// TIA Portal project "FactoryIO_Template_S7-1200_V15_V16" (V16)
// Vorlageprojekt für das Buch mit Zielsystem S7-1200

(* hardware
DEVICE "S7-1200-Station_1"  S7-1200 Station
   slot 0: "Baugruppenträger_0"  Rack  V1.0
   slot 1: "PLC_1"  CPU 1212C AC/DC/Rly  6ES7 212-1BE40-0XB0  V4.4
DEVICE "HMI_1"  KTP700 Basic PN
   slot 0: "HMI_1"  KTP700 Basic PN  6AV2 123-2GB03-0AX0  16.0.0.0
   slot 1: "HMI_RT_1"  KTP700 Basic PN  6AV2 123-2GB03-0AX0  16.0.0.0
   slot 5: "HMI_1.IE_CP_1"  PROFINET Interface  16.0.0.0
      slot 1: "PROFINET Interface_1"  PROFINET Interface
         slot 1: "Port_1"  Port
*)

// ===== PLC "PLC_1"  CPU 1212C AC/DC/Rly =====

VAR_GLOBAL   // PLC tag table "Standard-Variablentabelle"
   "SENSOR NIVEL" AT %IW30 : Int;
   "SENSOR CAUDAL" AT %IW32 : Int;
   "VALVULA LLENADO" AT %QW30 : Int;
   "VALVULA DESCARGA" AT %QW32 : Int;
   "VALOR CONSIGNA" AT %MD0 : DWord;
   "VISOR CONSIGNA" AT %QW34 : Int;
   "VISOR VALOR PROCESO" AT %QW36 : Int;
   "SET POINT" AT %IW34 : Int;
   "VALOR PROCESO" AT %MD12 : Real;
   "MARCA REAL SET  POINT mm" AT %MD4 : Real;
   "MARCA REAL VALOR PROCESO mm" AT %MD16 : Real;
   "MARCA REAL SET POINT %" AT %MD8 : Real;
   "VALOR MARCA REAL PROCESO %" AT %MD20 : Real;
   "START HMI" AT %M25.0 : Bool;
   "STOP HMI" AT %M26.0 : Bool;
   "INICIO" AT %M27.0 : Bool;
   "Start" AT %I0.0 : Bool;
   "Stop" AT %I0.2 : Bool;
   "INDICADOR 1" AT %Q0.0 : Bool;
   "INDICADOR 2" AT %Q0.2 : Bool;
   "ALTO" AT %M28.0 : Bool;
   "BAJO" AT %M29.0 : Bool;
   "PROCESO VALVULA LLENADO" AT %MD44 : Real;
   "VALVULA LLENADO %" AT %MD48 : Real;
   "ABRIR VALVULA" AT %M41.0 : Bool;
   "AUX SALIDA PID" AT %MD52 : Real;
   "AUX PID PROCESO" AT %MD56 : Real;
   "REGISTRO ACTIVO" AT %M60.0 : Bool;
   "PRIMER REGISTRO" AT %M64.0 : Bool;
   "NIVEL MAXIMO" AT %MD68 : Real;
   "NIVEL MINIMO" AT %MD72 : Real;
   "RESETEO" AT %M76.0 : Bool;
END_VAR

FUNCTION "MHJ-PLC-Lab-Function-S71200" : Void   // FC9000, SCL
{ S7_Optimized_Access := 'TRUE' }
VERSION : 0.1
   VAR_TEMP
      rdTimeReturn : Int;
      outputTime : DTL;
      SyncVal : Byte;
      forVal : Int;
      forVal_2 : Int;
      Value : Byte;
   END_VAR
   VAR CONSTANT
      CompVal : Byte := 16#34;
      Value_01 : Byte := 16#11;
      Value_01_DW : DWord := 16#A165_D992;
      Value_02_DW : DWord := 16#58BE_4401;
   END_VAR
BEGIN

   #Value:=PEEK(area := 16#82,
        dbNumber := 0,
        byteOffset := 511);
   #Value := #Value + 1;

   POKE(area := 16#82,
        dbNumber := 0,
        byteOffset := 511,
        value := #Value);

   POKE(area:=16#81,
        dbNumber:=0,
        byteOffset:=1016,
        value:=#Value_01_DW);
   POKE(area := 16#81,
        dbNumber := 0,
        byteOffset := 1020,
        value := #Value_02_DW);

   POKE(area := 16#81,
        dbNumber := 0,
        byteOffset := 511,
        value := B#16#00);

   FOR #forVal := 0 TO 120 DO
       FOR #forVal_2:=0 TO 10 DO
           #rdTimeReturn:=RD_SYS_T(#outputTime);
           #rdTimeReturn := WR_SYS_T(#outputTime);
           #rdTimeReturn := RD_SYS_T(#outputTime);
           #rdTimeReturn := WR_SYS_T(#outputTime);
       END_FOR;
       #SyncVal:= PEEK(area := 16#81,
                      dbNumber := 0,
                      byteOffset := 511);
       IF #SyncVal = #CompVal THEN
          GOTO M_1;
       END_IF;
   END_FOR;
   RETURN;

   M_1:
   POKE(area := 16#81,
        dbNumber := 0,
        byteOffset := 511,
        value := B#16#0);
END_FUNCTION

ORGANIZATION_BLOCK "Main"   // OB1, LAD, ProgramCycle
TITLE = "Main Program Sweep (Cycle)"
{ S7_Optimized_Access := 'TRUE' }
VERSION : 0.1
   VAR_INPUT
      Initial_Call : Bool;   // Initial call of this OB
      Remanence : Bool;   // =True, if remanent data are available
   END_VAR
BEGIN

REGION Network 1: Konnektierungsbaustein für PLC-Lab / CONEXION FACTORY IO
   // Im Netzwerk 1 wird der Konnektierungsbaustein für PLC-Lab aufgerufen.
   // Dieser Aufruf darf nicht entfernt werden!
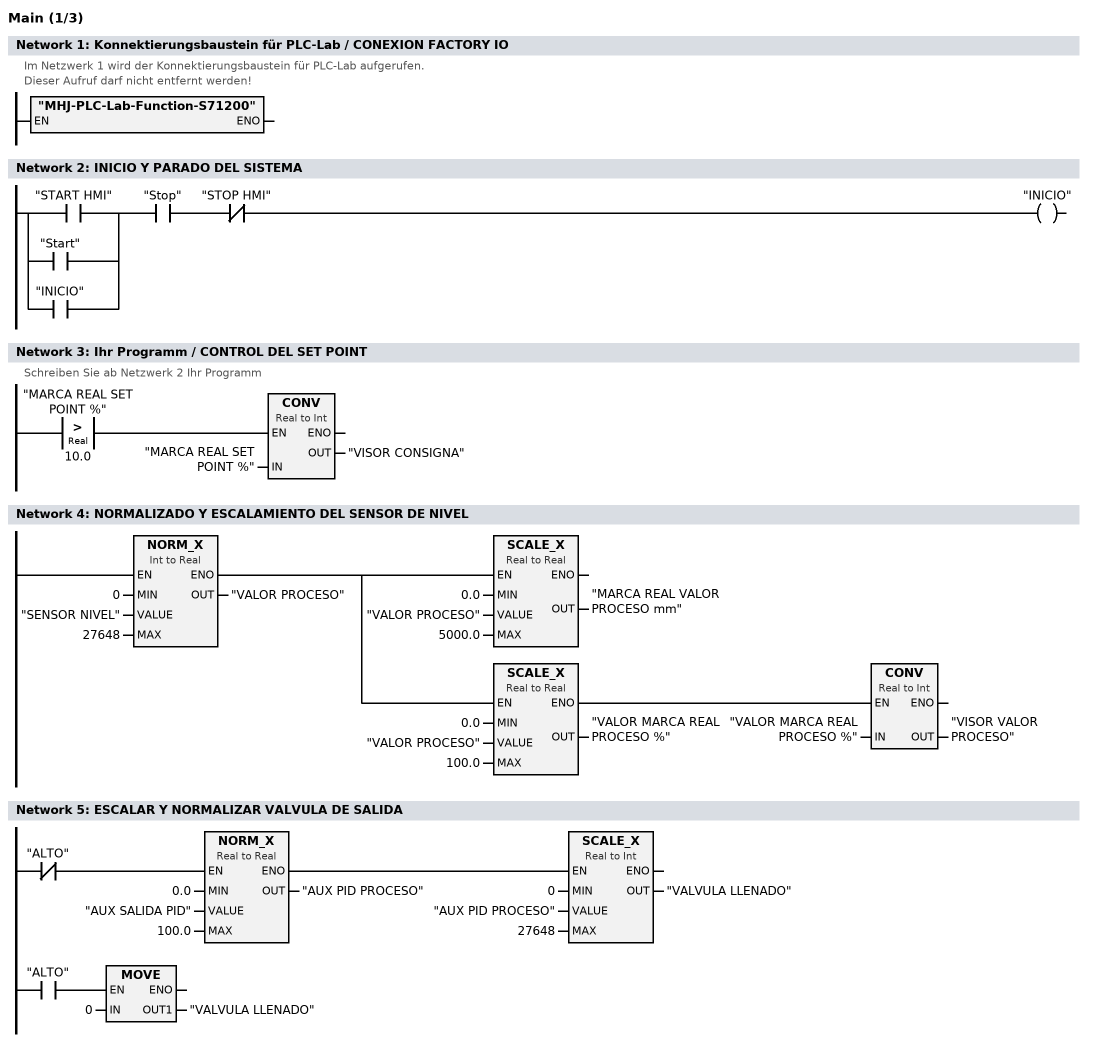
   RUNG wire#powerrail
      "MHJ-PLC-Lab-Function-S71200"()
   END_RUNG
   // the same network as SCL:
   "MHJ-PLC-Lab-Function-S71200"();
END_REGION

REGION Network 2: INICIO Y PARADO DEL SISTEMA
   RUNG wire#powerrail
      Contact( "START HMI" )
      wire#w1
      Contact( "Stop" )
      I_Contact( "STOP HMI" )
      Coil( "INICIO" )
   END_RUNG
   RUNG wire#powerrail
      Contact( "Start" )
   END_RUNG wire#w1
   RUNG wire#powerrail
      Contact( "INICIO" )
   END_RUNG wire#w1
   // the same network as SCL:
   "INICIO" := ("START HMI" OR "Start" OR "INICIO") AND "Stop" AND NOT "STOP HMI";
END_REGION

REGION Network 3: Ihr Programm / CONTROL DEL SET POINT
   // Schreiben Sie ab Netzwerk 2 Ihr Programm
   RUNG wire#powerrail
      { S7_Templates := "SrcType := Real" } GT_Contact(in1 := "MARCA REAL SET POINT %", in2 := 10.0)
      { S7_Templates := "[SrcType := Real, DestType := Int]" } Convert(in := "MARCA REAL SET POINT %", out => "VISOR CONSIGNA")
   END_RUNG
   // the same network as SCL:
   IF "MARCA REAL SET POINT %" > 10.0 THEN "VISOR CONSIGNA" := REAL_TO_INT("MARCA REAL SET POINT %"); END_IF;
END_REGION

REGION Network 4: NORMALIZADO Y ESCALAMIENTO DEL SENSOR DE NIVEL
   RUNG wire#powerrail
      { S7_Templates := "[SrcType := Int, DestType := Real]" } Normalize(min := 0, value := "SENSOR NIVEL", max := 27648, out => "VALOR PROCESO")
      wire#w1
      { S7_Templates := "[SrcType := Real, DestType := Real]" } Scale(min := 0.0, value := "VALOR PROCESO", max := 5000.0, out => "MARCA REAL VALOR PROCESO mm")
   END_RUNG
   RUNG wire#w1
      { S7_Templates := "[SrcType := Real, DestType := Real]" } Scale(min := 0.0, value := "VALOR PROCESO", max := 100.0, out => "VALOR MARCA REAL PROCESO %")
      { S7_Templates := "[SrcType := Real, DestType := Int]" } Convert(in := "VALOR MARCA REAL PROCESO %", out => "VISOR VALOR PROCESO")
   END_RUNG
   // the same network as SCL:
   "VALOR PROCESO" := NORM_X(MIN := 0, VALUE := "SENSOR NIVEL", MAX := 27648);
   "MARCA REAL VALOR PROCESO mm" := SCALE_X(MIN := 0.0, VALUE := "VALOR PROCESO", MAX := 5000.0);
   "VALOR MARCA REAL PROCESO %" := SCALE_X(MIN := 0.0, VALUE := "VALOR PROCESO", MAX := 100.0);
   "VISOR VALOR PROCESO" := REAL_TO_INT("VALOR MARCA REAL PROCESO %");
END_REGION

REGION Network 5: ESCALAR Y NORMALIZAR VALVULA DE SALIDA
   RUNG wire#powerrail
      I_Contact( "ALTO" )
      { S7_Templates := "[SrcType := Real, DestType := Real]" } Normalize(min := 0.0, value := "AUX SALIDA PID", max := 100.0, out => "AUX PID PROCESO")
      { S7_Templates := "[SrcType := Real, DestType := Int]" } Scale(min := 0, value := "AUX PID PROCESO", max := 27648, out => "VALVULA LLENADO")
   END_RUNG
   RUNG wire#powerrail
      Contact( "ALTO" )
      Move(in := 0, out1 => "VALVULA LLENADO")
   END_RUNG
   // the same network as SCL:
   IF NOT "ALTO" THEN
       "AUX PID PROCESO" := NORM_X(MIN := 0.0, VALUE := "AUX SALIDA PID", MAX := 100.0);
       "VALVULA LLENADO" := SCALE_X(MIN := 0, VALUE := "AUX PID PROCESO", MAX := 27648);
   END_IF;
   IF "ALTO" THEN "VALVULA LLENADO" := 0; END_IF;
END_REGION

REGION Network 6: ALARMAS DE NIVEL
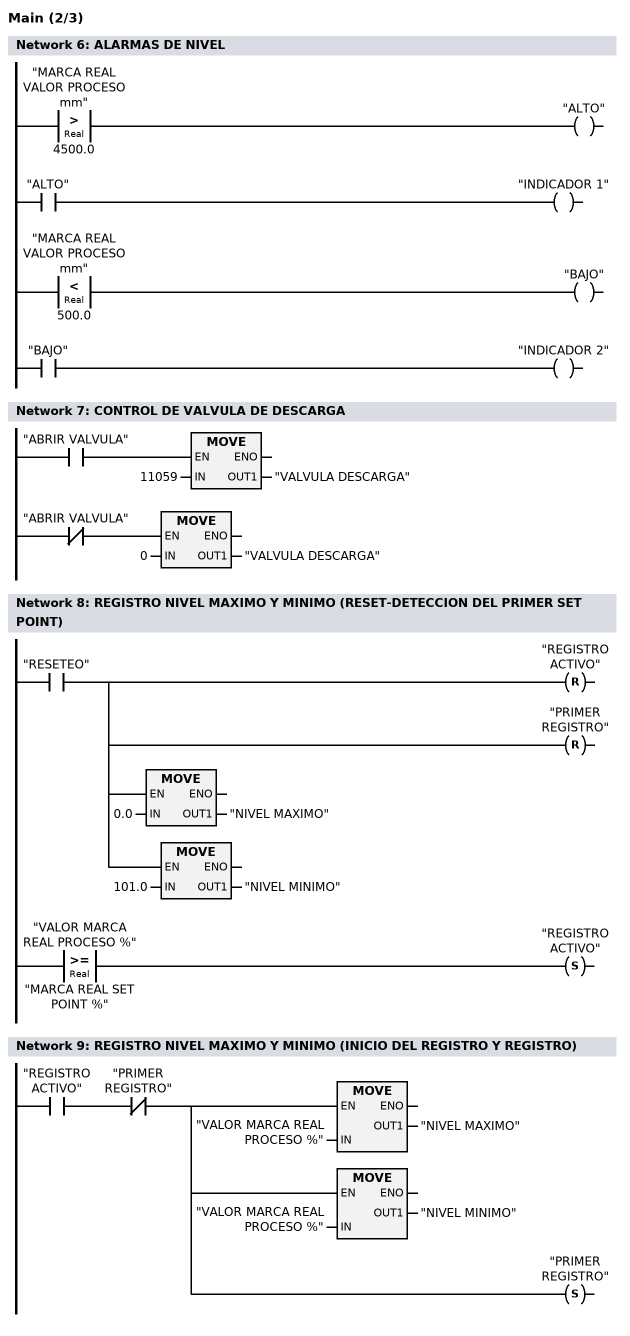
   RUNG wire#powerrail
      { S7_Templates := "SrcType := Real" } GT_Contact(in1 := "MARCA REAL VALOR PROCESO mm", in2 := 4500.0)
      Coil( "ALTO" )
   END_RUNG
   RUNG wire#powerrail
      Contact( "ALTO" )
      Coil( "INDICADOR 1" )
   END_RUNG
   RUNG wire#powerrail
      { S7_Templates := "SrcType := Real" } LT_Contact(in1 := "MARCA REAL VALOR PROCESO mm", in2 := 500.0)
      Coil( "BAJO" )
   END_RUNG
   RUNG wire#powerrail
      Contact( "BAJO" )
      Coil( "INDICADOR 2" )
   END_RUNG
   // the same network as SCL:
   "ALTO" := "MARCA REAL VALOR PROCESO mm" > 4500.0;
   "INDICADOR 1" := "ALTO";
   "BAJO" := "MARCA REAL VALOR PROCESO mm" < 500.0;
   "INDICADOR 2" := "BAJO";
END_REGION

REGION Network 7: CONTROL DE VALVULA DE DESCARGA
   RUNG wire#powerrail
      Contact( "ABRIR VALVULA" )
      Move(in := 11059, out1 => "VALVULA DESCARGA")
   END_RUNG
   RUNG wire#powerrail
      I_Contact( "ABRIR VALVULA" )
      Move(in := 0, out1 => "VALVULA DESCARGA")
   END_RUNG
   // the same network as SCL:
   IF "ABRIR VALVULA" THEN "VALVULA DESCARGA" := 11059; END_IF;
   IF NOT "ABRIR VALVULA" THEN "VALVULA DESCARGA" := 0; END_IF;
END_REGION

REGION Network 8: REGISTRO NIVEL MAXIMO Y MINIMO (RESET-DETECCION DEL PRIMER SET POINT)
   RUNG wire#powerrail
      Contact( "RESETEO" )
      wire#w1
      R_Coil( "REGISTRO ACTIVO" )
   END_RUNG
   RUNG wire#w1
      R_Coil( "PRIMER REGISTRO" )
   END_RUNG
   RUNG wire#w1
      Move(in := 0.0, out1 => "NIVEL MAXIMO")
   END_RUNG
   RUNG wire#w1
      Move(in := 101.0, out1 => "NIVEL MINIMO")
   END_RUNG
   RUNG wire#powerrail
      { S7_Templates := "SrcType := Real" } GE_Contact(in1 := "VALOR MARCA REAL PROCESO %", in2 := "MARCA REAL SET POINT %")
      S_Coil( "REGISTRO ACTIVO" )
   END_RUNG
   // the same network as SCL:
   IF "RESETEO" THEN
       "REGISTRO ACTIVO" := FALSE;
       "PRIMER REGISTRO" := FALSE;
       "NIVEL MAXIMO" := 0.0;
       "NIVEL MINIMO" := 101.0;
   END_IF;
   IF "VALOR MARCA REAL PROCESO %" >= "MARCA REAL SET POINT %" THEN "REGISTRO ACTIVO" := TRUE; END_IF;
END_REGION

REGION Network 9: REGISTRO NIVEL MAXIMO Y MINIMO (INICIO DEL REGISTRO Y REGISTRO)
   RUNG wire#powerrail
      Contact( "REGISTRO ACTIVO" )
      I_Contact( "PRIMER REGISTRO" )
      wire#w1
      Move(in := "VALOR MARCA REAL PROCESO %", out1 => "NIVEL MAXIMO")
   END_RUNG
   RUNG wire#w1
      Move(in := "VALOR MARCA REAL PROCESO %", out1 => "NIVEL MINIMO")
   END_RUNG
   RUNG wire#w1
      S_Coil( "PRIMER REGISTRO" )
   END_RUNG
   // the same network as SCL:
   IF "REGISTRO ACTIVO" AND NOT "PRIMER REGISTRO" THEN
       "NIVEL MAXIMO" := "VALOR MARCA REAL PROCESO %";
       "NIVEL MINIMO" := "VALOR MARCA REAL PROCESO %";
       "PRIMER REGISTRO" := TRUE;
   END_IF;
END_REGION

REGION Network 10: LOGICA DE REGISTRO DE MAXIMO Y MINIMOS
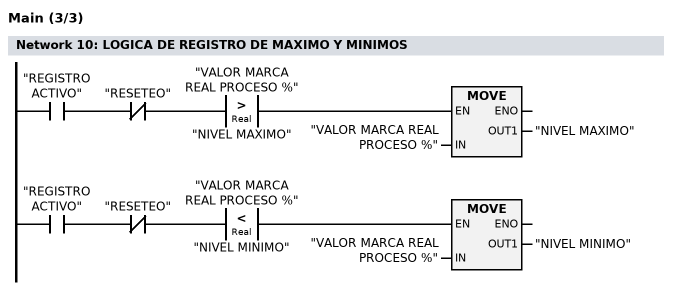
   RUNG wire#powerrail
      Contact( "REGISTRO ACTIVO" )
      I_Contact( "RESETEO" )
      { S7_Templates := "SrcType := Real" } GT_Contact(in1 := "VALOR MARCA REAL PROCESO %", in2 := "NIVEL MAXIMO")
      Move(in := "VALOR MARCA REAL PROCESO %", out1 => "NIVEL MAXIMO")
   END_RUNG
   RUNG wire#powerrail
      Contact( "REGISTRO ACTIVO" )
      I_Contact( "RESETEO" )
      { S7_Templates := "SrcType := Real" } LT_Contact(in1 := "VALOR MARCA REAL PROCESO %", in2 := "NIVEL MINIMO")
      Move(in := "VALOR MARCA REAL PROCESO %", out1 => "NIVEL MINIMO")
   END_RUNG
   // the same network as SCL:
   IF "REGISTRO ACTIVO" AND NOT "RESETEO" AND ("VALOR MARCA REAL PROCESO %" > "NIVEL MAXIMO") THEN
       "NIVEL MAXIMO" := "VALOR MARCA REAL PROCESO %";
   END_IF;
   IF "REGISTRO ACTIVO" AND NOT "RESETEO" AND ("VALOR MARCA REAL PROCESO %" < "NIVEL MINIMO") THEN
       "NIVEL MINIMO" := "VALOR MARCA REAL PROCESO %";
   END_IF;
END_REGION
END_ORGANIZATION_BLOCK

ORGANIZATION_BLOCK "Cyclic interrupt"   // OB30, LAD, CyclicInterrupt
{ S7_Optimized_Access := 'TRUE' }
VERSION : 0.1
   VAR_INPUT
      Initial_Call : Bool;   // Initial call of this OB
      Event_Count : Int;   // Events discarded
   END_VAR
BEGIN

REGION Network 1: PROCESO PID
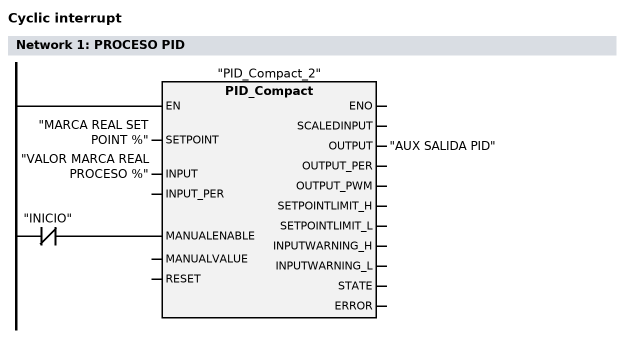
   "PID_Compact_2"(Setpoint := "MARCA REAL SET POINT %",   // PID_Compact
                   Input := "VALOR MARCA REAL PROCESO %",
                   ManualEnable := NOT "INICIO",
                   Output => "AUX SALIDA PID");
END_REGION
END_ORGANIZATION_BLOCK

(* ===== HMI "HMI_RT_1" =====
system functions are stored by id; their names below are inferred from use
connection "HMI_Connection_1": ETHERNET, SMART_S7_1200_OMS

HMI tags "Default tag table"
   "Tag_ScreenNumber" : UInt, internal
   "START HMI" : Bool = PLC "START HMI" AT %M25.0, 1 s
   "STOP HMI" : Bool = PLC "STOP HMI" AT %M26.0, 1 s
   "VALOR MARCA REAL PROCESO %" : Real = PLC "VALOR MARCA REAL PROCESO %" AT %MD20, 1 s
   "MARCA REAL SET POINT %" : Real = PLC "MARCA REAL SET POINT %" AT %MD8, 1 s
   "VALVULA LLENADO" : Int = PLC "VALVULA LLENADO" AT %QW30, 1 s
   "ALTO" : Bool = PLC ALTO AT %M28.0, 1 s
   "BAJO" : Bool = PLC BAJO AT %M29.0, 1 s
   "ABRIR VALVULA" : Bool = PLC "ABRIR VALVULA" AT %M41.0, 1 s
   "VALVULA LLENADO PROCESO %" : Real = PLC "VALVULA LLENADO %" AT %MD48, 1 s
   "AUX SALIDA PID" : Real = PLC "AUX SALIDA PID" AT %MD52, 1 s
   "NIVEL MAXIMO" : Real = PLC "NIVEL MAXIMO" AT %MD68, 1 s
   "NIVEL MINIMO" : Real = PLC "NIVEL MINIMO" AT %MD72, 1 s
   "RESETEO" : Bool = PLC RESETEO AT %M76.0, 1 s

Template "Template_1" 800x480
   Button "Exit" at 714,429 size 71x50; TextOff 'Exit'; PictureOff "ExitRuntime_KTP700_Basic_PN_TR"; PictureOn "ExitRuntime_KTP700_Basic_PN_TR"
      on Release: StopRuntime(0)
   Button "Template_Button" at 614,429 size 71x50; TextOff 'Text'
   Button "Template_Button_1" at 514,429 size 71x50; TextOff 'Text'
   Button "Template_Button_2" at 414,429 size 71x50; TextOff 'Text'
   Button "Template_Button_3" at 314,429 size 71x50; TextOff 'Text'
   Button "Template_Button_4" at 214,429 size 71x50; TextOff 'Text'
   Button "Start screen" at 114,429 size 71x50; TextOff 'Start screen'; PictureOff "NavigateHome_KTP700_Basic_PN_TR"; PictureOn "NavigateHome_KTP700_Basic_PN_TR"
      on Release: ActivateScreen("Root screen", 0)
   Button "Alarms" at 14,429 size 71x50; TextOff 'Alarms'; PictureOff "AlarmDisplay_KTP700_Basic_PN_TR"; PictureOn "AlarmDisplay_KTP700_Basic_PN_TR"
      on Release: function_ef3f5d25("Alarm window_Unacknowledged", -1)
   SymbolicIOField "Symbolic_IO_Field_Screen" at 93,9 size 600x33; TextOff '0'; TextOn '1'; TextList "TextList_ScreenNames"
      ProcessValue <- "Tag_ScreenNumber"
      on Change: ActivateScreenByNumber("Tag_ScreenNumber", 0)
   DateTimeField "HmiScreenItemData" at 695,25 size 105x25
   DateTimeField "HmiScreenItemData_1" at 695,0 size 105x25
   GraphicView "Logo" at 0,0 size 91x51; Picture "Logo of HMI_1"

screen "Root screen" 800x480, template "Template_1"
   on GenerateScreen: SetTag("Tag_ScreenNumber", 1)
   GraphicView "Graphic view_7" at 653,349 size 67x59; Picture "Graphic_6"
   TextField "HmiScreenItemData" at 227,49 size 397x25; Text 'CONTROL PID DE NIVEL DE TANQUE'
   Button "Button_2" at 41,212 size 144x52; TextOff 'STOP'
      on Press: SetBit("STOP HMI")
      on Release: ResetBit("STOP HMI")
   Button "Button_1" at 41,128 size 144x52; TextOff 'START'
      on Press: SetBit("START HMI")
      on Release: ResetBit("START HMI")
   GraphicView "Graphic view_1" at 609,145 size 170x211; Picture "Graphic_1"
   Bar "Bar_1" at 635,165 size 116x164; MinimumValue 0; MaximumValue 100
      ProcessValue <- "VALOR MARCA REAL PROCESO %"
   GraphicView "Graphic view_2" at 616,80 size 50x58; Picture "Graphic_3"
   GraphicView "Graphic view_3" at 611,331 size 46x64; Picture "Graphic_3"
   GraphicView "Graphic view_4" at 655,86 size 59x66; Picture "Graphic_4"
   TextField "Text field_1" at 667,85 size 107x23; Text 'V. LLENADO'
   TextField "Text field_2" at 684,377 size 103x23; Text 'V. VACIADO'
   IOField "I/O field_1" at 268,232 size 96x32; FormatPattern s999999999.999
      ProcessValue <- "VALOR MARCA REAL PROCESO %"
   IOField "I/O field_2" at 264,155 size 96x32; FormatPattern s999999999.999
      ProcessValue <- "MARCA REAL SET POINT %"
   TextField "Text field_3" at 264,126 size 94x23; Text 'SET POINT'
   Circle "Circle_1" at 467,322 size 37x37
      Appearance <- "ALTO"
   TextField "Text field_4" at 256,207 size 126x23; Text 'NIVEL ACTUAL'
   TextField "Text field_5" at 264,283 size 102x23; Text 'SALIDA PID'
   Circle "Circle_3" at 531,322 size 37x37
      Appearance <- "BAJO"
   TextField "Text field_6" at 459,302 size 57x23; Text 'LLENO'
   TextField "Text field_7" at 519,302 size 63x23; Text 'VACIO'
   Switch "Switch_1" at 60,318 size 93x39; CaptionText 'Switch'; TextOff 'OFF'; TextOn 'ON'
      on SwitchOn: SetBit("ABRIR VALVULA")
      on SwitchOff: ResetBit("ABRIR VALVULA")
   TextField "Text field_9" at 24,282 size 174x23; Text 'VACIAR CONTENIDO'
   IOField "I/O field_3" at 268,316 size 96x32; FormatPattern s999999999.999
      ProcessValue <- "AUX SALIDA PID"
   IOField "I/O field_4" at 463,150 size 96x32; FormatPattern s999999999.999
      ProcessValue <- "NIVEL MAXIMO"
   IOField "I/O field_5" at 462,212 size 96x32; FormatPattern s999999999.999
      ProcessValue <- "NIVEL MINIMO"
   TextField "Text field_8" at 450,186 size 119x23; Text 'MENOR NIVEL'
   TextField "Text field_10" at 455,124 size 120x23; Text 'MAYOR NIVEL'
   Button "Button_3" at 464,256 size 96x32; TextOff 'RESET'
      on Press: SetBit("RESETEO")
      on Release: ResetBit("RESETEO")
*)